Fanuc KAREL source: ko00108.KL

-- PROVISIONAL review KL for V1013-1; original PC SHA256 48f30c1fd32adf7a70428de5d2d4f435ce2cfbd46525c24076fc656b885cf3ed
-- Incomplete behavior may be omitted. Consult companion uncertainty JSON. Do not deploy.
PROGRAM KO00108
%NOLOCKGROUP
VAR
  A : REAL
  B : REAL
  OUT : REAL
BEGIN
  -- UNRESOLVED_PC offsets 5-13; opcodes 9D,64,23
  -- UNRESOLVED_PC offsets 18-30; opcodes 2E,64,23
  -- UNRESOLVED_PC offsets 35-56; opcodes 27,22,22,76,23
  -- UNRESOLVED_PC offsets 61-65; opcodes 7F
END KO00108
